Fanuc KAREL source: KT00741.KL

PROGRAM KT00741
%NOLOCKGROUP
VAR
  ARG: ARRAY[4] OF SHORT
  OUT: INTEGER
BEGIN
  OUT = ARRAY_LEN(ARG)
END KT00741
